(* IEC 61131-3 sources: plc-process-lib/tests/POUs/Helpers/FB_TestDevice, 7 files *)

(* ---- FB_TestDevice.decl.st ---- *)
// Назначение: тестовое устройство — наследник FB_DeviceBase, на котором проверяется база.
//             Тело — нормативный порядок цикла устройства (docs/fb/FB_DeviceBase.md): ResolveTime
//             до вложенного FB_Delay, BeginCycle, AcceptCfg(CheckConfig) с LKG, Reset с
//             фиксируемым отказом, ProcessMode, команды пуск/стоп (SwitchRemoteMode при «Стоп» в
//             Auto), безопасный выход, RunAlarms, FinishCycle. Переопределяет хук OnModeChanged
//             (безударность, снятие отказа при входе в OutOfService) и записывает его вызовы.
//             xInputLike = TRUE ведёт себя как AI/DI: режим в stModeMem, Manual = CheckFunction.
//             Только для тестов.
// Автор:      kr0nsch
// Версия:     0.1.0
// Документ:   docs/TESTING.md, раздел «Тестовое устройство»
FUNCTION_BLOCK FB_TestDevice EXTENDS FB_DeviceBase
VAR CONSTANT
    CFG_GAIN   : WORD := 16#0001;  // wCfgErr бит 0: rGain не конечен или <= 0
    CFG_ALARM  : WORD := 16#0002;  // wCfgErr бит 1: приоритет тревоги вне перечисления (CheckAlarmCfg)
    STS_OUTPUT : WORD := 16#0001;  // wStatus бит 0: выход включён
    STS_FAULT  : WORD := 16#0002;  // wStatus бит 1: зафиксирован отказ
    FLT_LATCH  : WORD := 16#0001;  // wFault бит 0: зафиксированный механический отказ
    GAIN_SCALE : REAL := 10.0;     // rOut_eu = rGain * GAIN_SCALE
END_VAR
VAR_INPUT
    xAutoRun        : BOOL;                                   // запрос автоматики «работать»
    xLocal          : BOOL;                                   // переключатель «Местное»
    xMoving         : BOOL;                                   // механизм в движении: вывод из работы запрещён
    xFaultCause     : BOOL;                                   // причина механического отказа (фиксируется)
    xShedToManual   : BOOL;                                   // логика устройства переводит в Manual
    xLocalSupported : BOOL := TRUE;                           // FALSE — как у AI/DI: режима Local нет
    xInputLike      : BOOL;                                   // TRUE — как AI/DI (задаётся до первого вызова)
    uiAlarmSlots    : UINT := 8;                              // используемых слотов (в первом вызове)
    eTypeSel        : E_DeviceType := E_DeviceType.Valve;     // тип для eDevType (в первом вызове)
    eDevStatusIn    : E_Ne107Status := E_Ne107Status.Good;    // вклад логики устройства в NE 107
    wWarnIn         : WORD;                                   // предупреждения устройства
    axCondIn        : ARRAY[0..GVL_Const.DEV_ALARMS_MAX - 1] OF BOOL;   // условия тревог слотов
    axSuppressIn    : ARRAY[0..GVL_Const.DEV_ALARMS_MAX - 1] OF BOOL;   // подавление по условию
    rValueIn        : REAL;                                   // значение процесса для событий
END_VAR
VAR_IN_OUT
    stCmd    : ST_TestDeviceCmd;   // команды
    stRetain : ST_DeviceRetain;    // энергонезависимые данные (при xInputLike не используются)
END_VAR
VAR_IN_OUT CONSTANT
    stCfg : ST_TestDeviceCfg;      // конфигурация
END_VAR
VAR_OUTPUT
    xOutput : BOOL;                // выход механизма; безопасное состояние — FALSE
    rOut_eu : REAL;                // значение по LKG: rGain * 10; 0 — корректной Cfg не было
    stSts   : ST_TestDeviceSts;    // состояние для HMI
END_VAR
VAR
    stCfgLkg       : ST_TestDeviceCfg;   // последняя корректная конфигурация (LKG)
    fbRunDelay     : FB_Delay;           // задержка включения в Auto — вызывается до BeginCycle
    xManualRun     : BOOL;               // ручная защёлка «работать»
    xFaultLatched  : BOOL;               // зафиксированный механический отказ
    xFaultAdd      : BOOL;               // точка расширения: доп. причина отказа (пишет наследник до SUPER^)
    uiBodyCalls    : UINT;               // сколько раз выполнено это тело
    ltDtSeen       : LTIME;              // ltDt последнего вызова (после BeginCycle)
    // --- журнал хука OnModeChanged ---
    uiHookCalls    : UINT;               // вызовов хука
    eHookOld       : E_DeviceMode := E_DeviceMode.Manual;   // eOld последнего вызова
    eHookNew       : E_DeviceMode := E_DeviceMode.Manual;   // eNew последнего вызова
    xHookInFirst   : BOOL;               // хук вызывался в первом вызове (xFirstCall = TRUE)
    udiHookTrace   : UDINT;              // порядок частей хука: цифра на уровень иерархии (1 — этот ФБ)
END_VAR
VAR_TEMP
    xResetNow : BOOL;                    // Reset в этом вызове
    eRes      : E_CmdResult;             // результат ProcessMode
    eDevSt    : E_Ne107Status;           // статус логики устройства
    uiLoop    : UINT;                    // номер слота + 1
    uiSlot    : UINT;                    // номер слота
END_VAR

(* ---- CheckConfig.method.decl.st ---- *)
// Проверка конфигурации: биты wCfgErr тестового устройства. Только считает, ничего не меняет
METHOD PROTECTED CheckConfig : WORD
VAR_IN_OUT CONSTANT
    stCfgIn : ST_TestDeviceCfg;   // проверяемая конфигурация
END_VAR
VAR
    wErr : WORD;                  // непройденные проверки
END_VAR

(* ---- CheckConfig.method.impl.st ---- *)
IF NOT F_IsFinite(rIn := stCfgIn.rGain) OR stCfgIn.rGain <= 0.0 THEN
    wErr := wErr OR CFG_GAIN;
END_IF
IF NOT CheckAlarmCfg(astCfg := stCfgIn.astAlarm) THEN
    wErr := wErr OR CFG_ALARM;
END_IF
CheckConfig := wErr;

(* ---- FB_TestDevice.impl.st ---- *)
// 0. Источник времени до BeginCycle: вложенный FB_Delay ниже вызывается раньше BeginCycle (как
//    fbVfdCommLoss у FB_MotorVfd, контракт 14.2); первый вызов — сразу с подменным временем
ResolveTime();
uiBodyCalls := uiBodyCalls + 1;
IF xFirstCall THEN
    uiAlarmCount := MIN(uiAlarmSlots, GVL_Const.DEV_ALARMS_MAX);
    eDevType := eTypeSel;
    xManualIsCheck := xInputLike;
    IF xInputLike THEN
        stModeMem.eRemoteMode := E_DeviceMode.Auto;
    ELSE
        stModeMem.eRemoteMode := E_DeviceMode.Manual;
    END_IF
END_IF
fbRunDelay(xIn := xAutoRun, tOnDelay := stCfgLkg.tRunDelay, itfTime := itfTimeAct);

// 1. Время
BeginCycle();
ltDtSeen := ltDt;

// 2. Конфигурация (LKG)
IF AcceptCfg(wErr := CheckConfig(stCfgIn := stCfg)) THEN
    stCfgLkg := stCfg;
END_IF

// 3. Reset: снимает зафиксированный отказ, если причина ушла
xResetNow := xResetReq OR stCmd.stCommon.xReset;
IF xResetNow THEN
    IF xFaultCause OR xFaultAdd THEN
        SetCmdResult(eResult := E_CmdResult.RejectedFault);
    ELSE
        xFaultLatched := FALSE;
        SetCmdResult(eResult := E_CmdResult.Accepted);
    END_IF
END_IF

// 4. Режим (AI/DI-подобное устройство — память режима stModeMem вместо stRetain)
IF xInputLike THEN
    eRes := ProcessMode(xLocalSel := xLocal, xLocalSupported := xLocalSupported, xOosAllowed := NOT xMoving,
                        stCmd := stCmd.stCommon, stRetain := stModeMem);
ELSE
    eRes := ProcessMode(xLocalSel := xLocal, xLocalSupported := xLocalSupported, xOosAllowed := NOT xMoving,
                        stCmd := stCmd.stCommon, stRetain := stRetain);
END_IF
IF eRes <> E_CmdResult.None THEN
    SetCmdResult(eResult := eRes);
END_IF

// 5. Команды устройства: xStop старше xStart; логика переводит в Manual (SwitchRemoteMode)
IF stCmd.xStop THEN
    IF eMode = E_DeviceMode.Auto OR eMode = E_DeviceMode.Manual THEN
        IF xInputLike THEN
            SwitchRemoteMode(eNew := E_DeviceMode.Manual, stRetain := stModeMem);
        ELSE
            SwitchRemoteMode(eNew := E_DeviceMode.Manual, stRetain := stRetain);
        END_IF
        xManualRun := FALSE;
        SetCmdResult(eResult := E_CmdResult.Accepted);
    ELSE
        SetCmdResult(eResult := E_CmdResult.RejectedMode);
    END_IF
ELSIF stCmd.xStart THEN
    IF eMode <> E_DeviceMode.Manual THEN
        SetCmdResult(eResult := E_CmdResult.RejectedMode);
    ELSIF NOT xCfgEverOk THEN
        SetCmdResult(eResult := E_CmdResult.RejectedCfg);
    ELSIF xFaultLatched OR xFaultCause OR xFaultAdd THEN
        SetCmdResult(eResult := E_CmdResult.RejectedFault);
    ELSE
        xManualRun := TRUE;
        SetCmdResult(eResult := E_CmdResult.Accepted);
    END_IF
END_IF
stCmd.xStart := FALSE;
stCmd.xStop := FALSE;
IF xShedToManual THEN
    IF xInputLike THEN
        SwitchRemoteMode(eNew := E_DeviceMode.Manual, stRetain := stModeMem);
    ELSE
        SwitchRemoteMode(eNew := E_DeviceMode.Manual, stRetain := stRetain);
    END_IF
END_IF

// 6. Логика по LKG. Отказ фиксируется вне OutOfService; безопасный выход — FALSE без корректной
//    Cfg и при отказе (ручная защёлка снимается)
IF (xFaultCause OR xFaultAdd) AND eMode <> E_DeviceMode.OutOfService THEN
    xFaultLatched := TRUE;
END_IF
IF NOT xCfgEverOk OR xFaultLatched THEN
    xOutput := FALSE;
    xManualRun := FALSE;
ELSIF eMode = E_DeviceMode.Auto THEN
    xOutput := fbRunDelay.xOut;
ELSIF eMode = E_DeviceMode.Manual THEN
    xOutput := xManualRun;
ELSE
    xOutput := FALSE;
END_IF
IF xCfgEverOk THEN
    rOut_eu := stCfgLkg.rGain * GAIN_SCALE;
ELSE
    rOut_eu := 0.0;
END_IF

// 7. Тревоги
FOR uiLoop := 1 TO GVL_Const.DEV_ALARMS_MAX DO
    uiSlot := uiLoop - 1;
    axAlmCond[uiSlot] := axCondIn[uiSlot];
    axAlmSuppress[uiSlot] := axSuppressIn[uiSlot];
    arAlmValue[uiSlot] := rValueIn;
END_FOR
RunAlarms(udiIdBase := stCfgLkg.udiAlarmIdBase, stCmd := stCmd.stCommon, astCfg := stCfgLkg.astAlarm);

// 8. Состояние
stSts.rOut_eu := rOut_eu;
IF xFaultLatched THEN
    eDevSt := E_Ne107Status.Failure;
ELSE
    eDevSt := eDevStatusIn;
END_IF
FinishCycle(eDevStatus := eDevSt,
            xAvailableDev := (eMode = E_DeviceMode.Auto) AND NOT xFaultLatched,
            wLow := SEL(xOutput, 0, STS_OUTPUT) OR SEL(xFaultLatched, 0, STS_FAULT),
            wFaultBits := SEL(xFaultLatched, 0, FLT_LATCH),
            wWarnBits := wWarnIn,
            stCommon := stSts.stCommon);

(* ---- OnModeChanged.method.decl.st ---- *)
// Хук смены режима: сначала база (SUPER^), затем запись вызова для тестов, безударность
// Auto → Manual (ручная защёлка := текущий выход) и снятие зафиксированного отказа при входе в
// OutOfService. VAR_IN_OUT устройства не трогает (R2)
METHOD PROTECTED OnModeChanged
VAR_INPUT
    eOld : E_DeviceMode;   // режим до смены
    eNew : E_DeviceMode;   // новый режим
END_VAR

(* ---- OnModeChanged.method.impl.st ---- *)
SUPER^.OnModeChanged(eOld := eOld, eNew := eNew);
uiHookCalls := uiHookCalls + 1;
eHookOld := eOld;
eHookNew := eNew;
xHookInFirst := xHookInFirst OR xFirstCall;
udiHookTrace := udiHookTrace * 10 + 1;
IF eOld = E_DeviceMode.Auto AND eNew = E_DeviceMode.Manual THEN
    xManualRun := xOutput;
END_IF
IF eNew = E_DeviceMode.OutOfService THEN
    xFaultLatched := FALSE;
END_IF

(* ---- ProbeAlarmCfg.method.decl.st ---- *)
// Открывает защищённый CheckAlarmCfg для тестов: проверка массива ST_AlarmCfg любой Cfg устройства
METHOD PUBLIC ProbeAlarmCfg : BOOL
VAR_IN_OUT CONSTANT
    astCfgIn : ARRAY[0..GVL_Const.DEV_ALARMS_MAX - 1] OF ST_AlarmCfg;   // проверяемый массив
END_VAR
